// SIMATIC S7-200 project (STEP 7-Micro/WIN), CPU 224XP CN REL 02.01

SYMBOL_TABLE USER1
Pos_Actual       VD100    // Posicion actual en cuentas (REAL)
Pos_Anterior     VD104    // Posicion ciclo anterior (REAL)
Vel_Actual       VD108    // Velocidad calculada en cuentas/s (REAL)
Setpoint         VD112    // Posicion objetivo en cuentas (REAL)
Accion_Control   VD116    // U calculada (con signo) (REAL)
K1               VD120    // Ganancia de posicion (97.26) (REAL)
K2               VD124    // Ganancia de velocidad (25.64) (REAL)
N                VD132    // Ganancia de pre-compensacion (REAL)
U_Abs            VD128    // Valor absoluto de la accion de control (REAL)
Seta_Emergencia  I1.4     // Entrada de seguridad (NC: 1=OK, 0=EMERGENCIA)
Variador_Run     Q0.0     // Mando Marcha/Paro (1=Run, 0=Stop)
Variador_Dir     Q0.1     // Mando Direccion (0=FWD, 1=REV)
Salida_Analog    AQW0     // Consigna de velocidad (0-32000)
INPUT            VD136    // Entrada manual para el setpoint
END_SYMBOL_TABLE

SYMBOL_TABLE S7-200 Symbols
Always_On        SM0.0    // Always ON
First_Scan_On    SM0.1    // ON for the first scan cycle only
Time_0_Intrvl    SMB34    // Specifies time interval (in 1-ms increments from 5 to 255) of interrupt 0.
HSC0_Ctrl        SMB37    // Configure and control HSC0
HSC0_CV          SMD38    // HSC0 new current value
HSC0_PV          SMD42    // HSC0 new preset value
END_SYMBOL_TABLE

ORGANIZATION_BLOCK MAIN:OB1
TITLE=
BEGIN
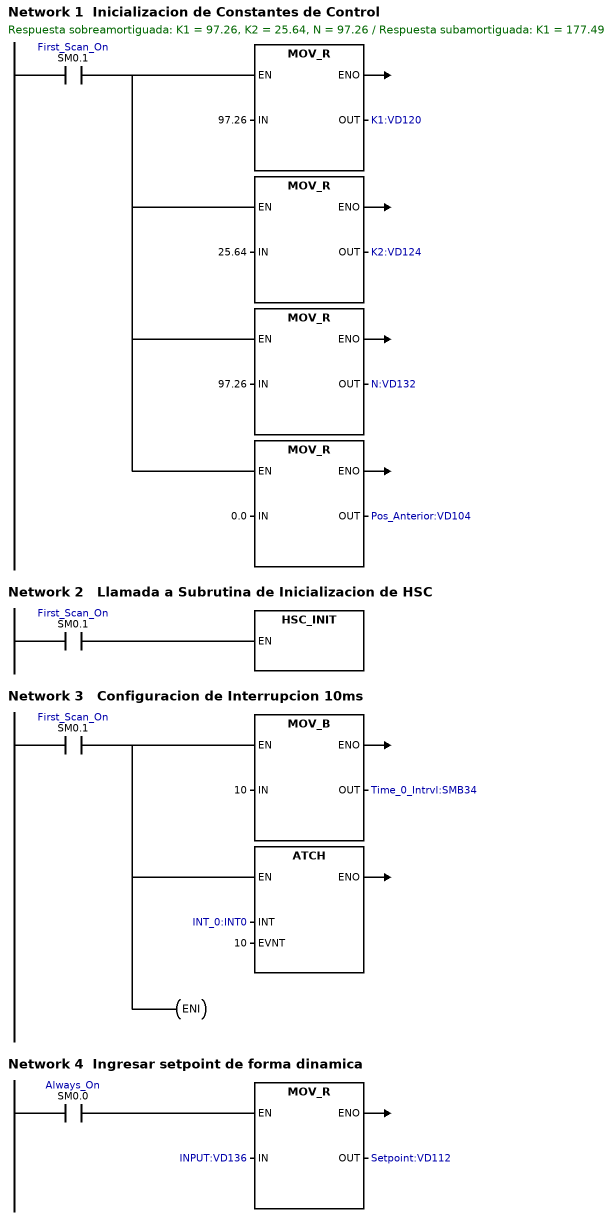
Network 1 // Inicializacion de Constantes de Control
// Respuesta sobreamortiguada: K1 = 97.26, K2 = 25.64, N = 97.26
// Respuesta subamortiguada: K1 = 177.49, K2 = 2.89, N = 177.49
// K1
// K2
// N (Pre-compensacion inicial = K1)
// Reset Pos_Anterior
LD     First_Scan_On:SM0.1
MOVR   97.26, K1:VD120
MOVR   25.64, K2:VD124
MOVR   97.26, N:VD132
MOVR   0.0, Pos_Anterior:VD104
Network 2 //  Llamada a Subrutina de Inicializacion de HSC
// Llamada a HSC_INIT
LD     First_Scan_On:SM0.1
CALL   HSC_INIT:SBR1
Network 3 //  Configuracion de Interrupcion 10ms
LD     First_Scan_On:SM0.1
MOVB   10, Time_0_Intrvl:SMB34
ATCH   INT_0:INT0, 10
ENI
Network 4 // Ingresar setpoint de forma dinamica
LD     Always_On:SM0.0
MOVR   INPUT:VD136, Setpoint:VD112
END_ORGANIZATION_BLOCK

SUBROUTINE_BLOCK HSC_INIT:SBR1
TITLE=
BEGIN
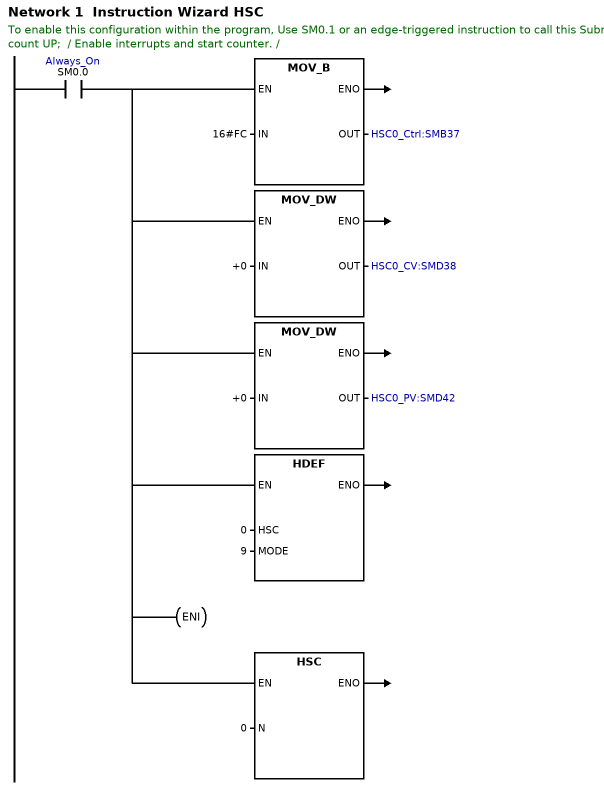
Network 1 // Instruction Wizard HSC
// To enable this configuration within the program, Use SM0.1 or an edge-triggered instruction to call this Subroutine once from the MAIN program block.  
// Configure HC0 for Mode 9; CV = 0; PV = 0; count UP; 
// Enable interrupts and start counter.
// 
//Set control bits: count UP; rate 1X; enabled; 
//Load CV
//Load PV
LD     Always_On:SM0.0
MOVB   16#FC, HSC0_Ctrl:SMB37
MOVD   +0, HSC0_CV:SMD38
MOVD   +0, HSC0_PV:SMD42
HDEF   0, 9
ENI
HSC    0
END_SUBROUTINE_BLOCK

INTERRUPT_BLOCK INT_0:INT0
TITLE=
BEGIN
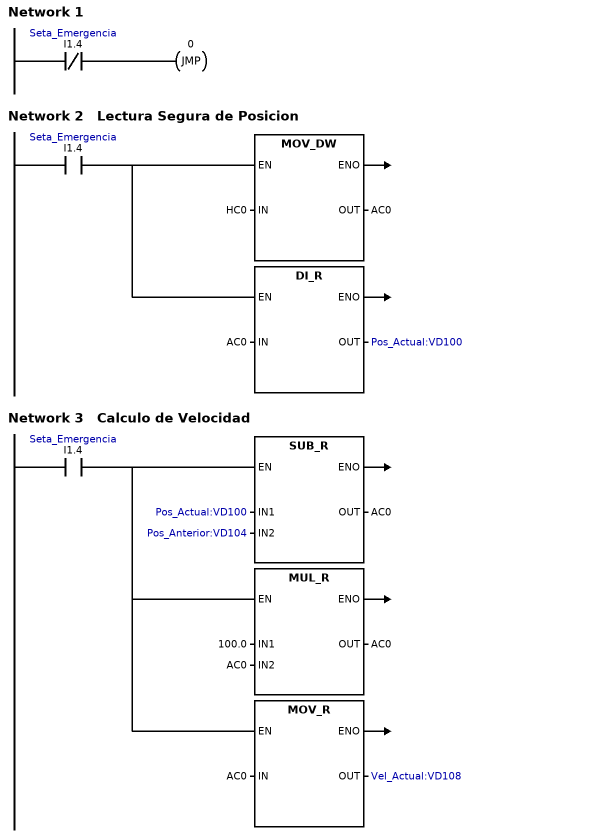
Network 1
LDN    Seta_Emergencia:I1.4
JMP    0
Network 2 //  Lectura Segura de Posicion
// Primero mover a AC0 (Búfer)
// Luego convertir a REAL
LD     Seta_Emergencia:I1.4
MOVD   HC0, AC0
DTR    AC0, Pos_Actual:VD100
Network 3 //  Calculo de Velocidad
// Delta Pos
// Equivalente a / 0.01s (Mas estable)
// VD108 = Vel_Actual
LD     Seta_Emergencia:I1.4
MOVR   Pos_Actual:VD100, AC0
-R     Pos_Anterior:VD104, AC0
*R     100.0, AC0
MOVR   AC0, Vel_Actual:VD108
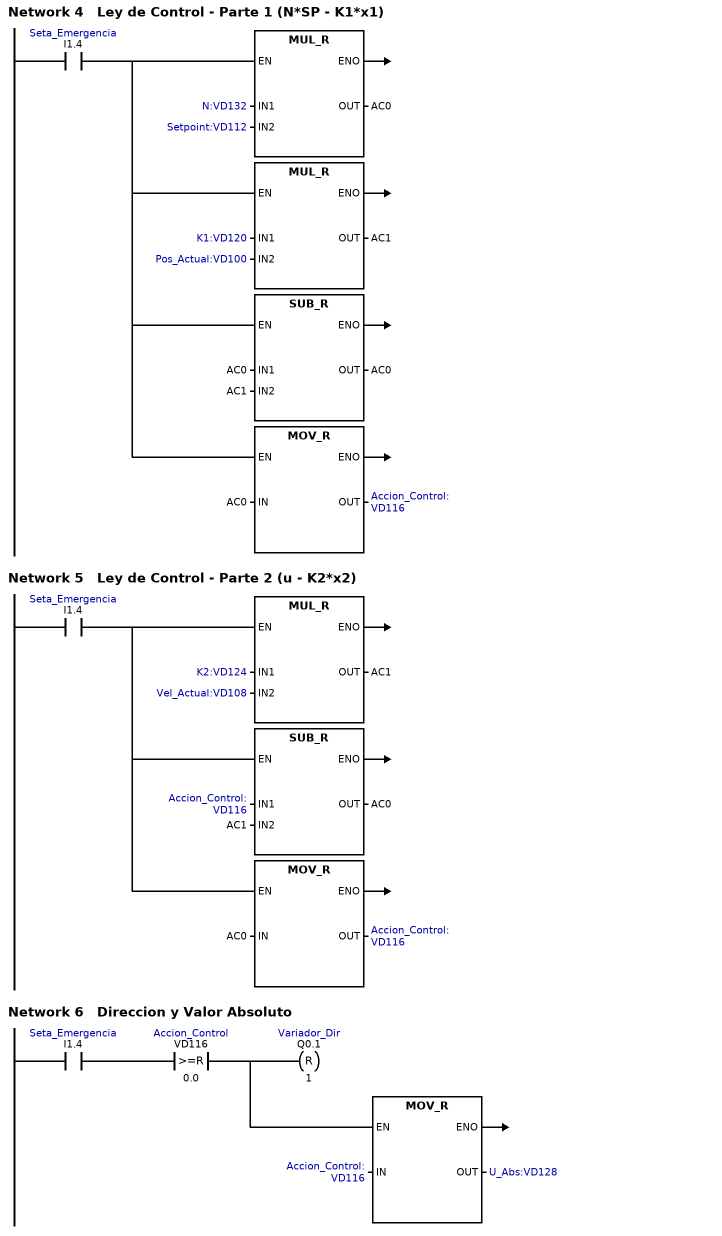
Network 4 //  Ley de Control - Parte 1 (N*SP - K1*x1)
// N
// N * SP
// K1
// K1 * x1
// AC0 = N*SP - K1*x1
// Guardado temporal
LD     Seta_Emergencia:I1.4
MOVR   N:VD132, AC0
*R     Setpoint:VD112, AC0
MOVR   K1:VD120, AC1
*R     Pos_Actual:VD100, AC1
-R     AC1, AC0
MOVR   AC0, Accion_Control:VD116
Network 5 //  Ley de Control - Parte 2 (u - K2*x2)
// K2
// K2 * x2
// AC0 = Accion Final
// Accion_Control final
LD     Seta_Emergencia:I1.4
MOVR   K2:VD124, AC1
*R     Vel_Actual:VD108, AC1
MOVR   Accion_Control:VD116, AC0
-R     AC1, AC0
MOVR   AC0, Accion_Control:VD116
Network 6 //  Direccion y Valor Absoluto
// FWD
LD     Seta_Emergencia:I1.4
AR>=   Accion_Control:VD116, 0.0
R      Variador_Dir:Q0.1, 1
MOVR   Accion_Control:VD116, U_Abs:VD128
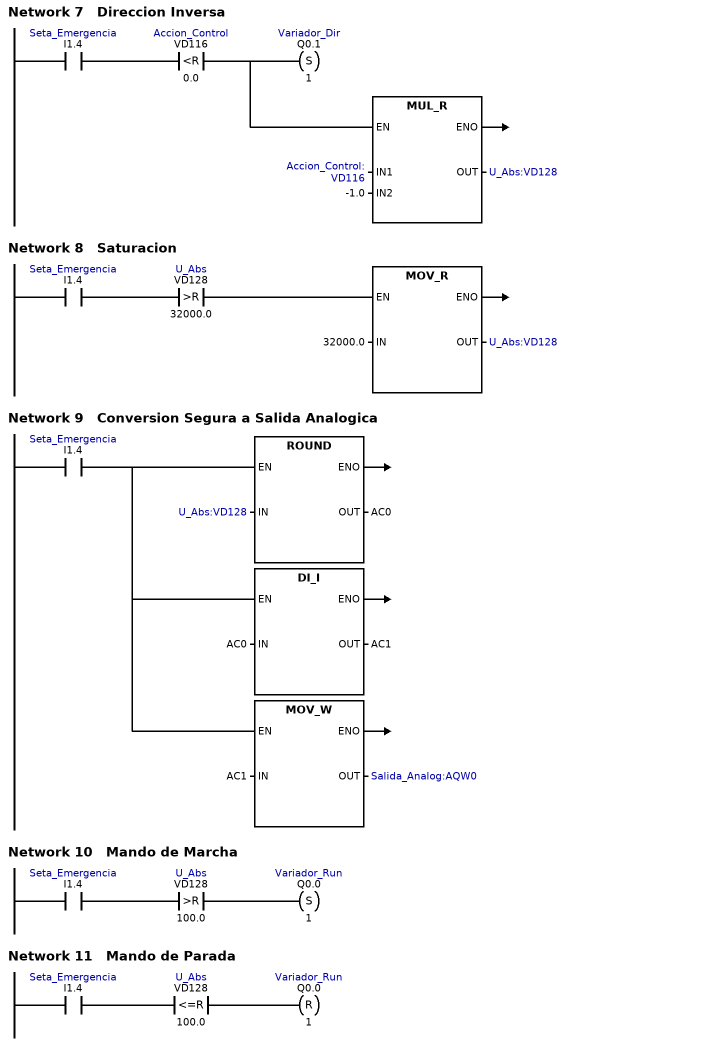
Network 7 //  Direccion Inversa
// REV
// |u|
LD     Seta_Emergencia:I1.4
AR<    Accion_Control:VD116, 0.0
S      Variador_Dir:Q0.1, 1
MOVR   Accion_Control:VD116, U_Abs:VD128
*R     -1.0, U_Abs:VD128
Network 8 //  Saturacion
LD     Seta_Emergencia:I1.4
AR>    U_Abs:VD128, 32000.0
MOVR   32000.0, U_Abs:VD128
Network 9 //  Conversion Segura a Salida Analogica
// Convertir a DINT en AC0
// Convertir DINT a INT en AC1 (Búfer)
// Mover Word a Salida (Forma mas segura)
LD     Seta_Emergencia:I1.4
ROUND  U_Abs:VD128, AC0
DTI    AC0, AC1
MOVW   AC1, Salida_Analog:AQW0
Network 10 //  Mando de Marcha
LD     Seta_Emergencia:I1.4
AR>    U_Abs:VD128, 100.0
S      Variador_Run:Q0.0, 1
Network 11 //  Mando de Parada
LD     Seta_Emergencia:I1.4
AR<=   U_Abs:VD128, 100.0
R      Variador_Run:Q0.0, 1
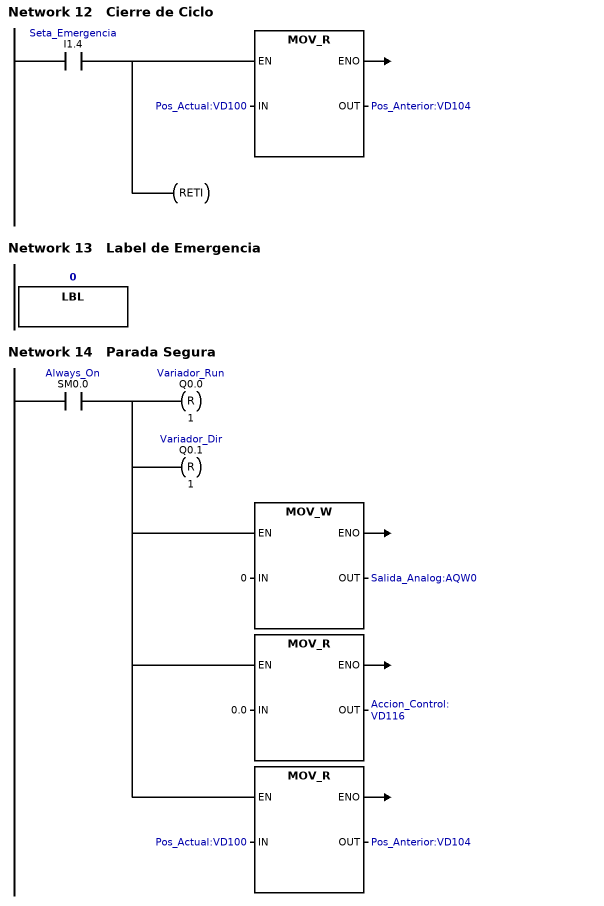
Network 12 //  Cierre de Ciclo
// Guardar Posicion para sig. ciclo
LD     Seta_Emergencia:I1.4
MOVR   Pos_Actual:VD100, Pos_Anterior:VD104
CRETI
Network 13 //  Label de Emergencia
LBL    0
Network 14 //  Parada Segura
LD     Always_On:SM0.0
R      Variador_Run:Q0.0, 1
R      Variador_Dir:Q0.1, 1
MOVW   0, Salida_Analog:AQW0
MOVR   0.0, Accion_Control:VD116
MOVR   Pos_Actual:VD100, Pos_Anterior:VD104
END_INTERRUPT_BLOCK
